(* IEC 61131-3 sources: rusty/compiler/plc_cfc/fixtures/blocks/valid/function_void, 1 file *)

(* ---- myVoid.st ---- *)
FUNCTION myVoid
VAR_INPUT
    in : DINT;
END_VAR
VAR_OUTPUT
    out : DINT;
END_VAR
    out := in * 2;
END_FUNCTION
